PROGRAM prg_Initialise
VAR_INPUT
	ResumeSFC       : BOOL; 		(*	not automatic	*)
	//Added SFC Cycle handle Variables
	
	SFCInit             : BOOL;  //shachar
END_VAR

VAR


(* 8888888888888888   SFC   8888888888888888888888*)
	sCycleName	        : STRING;
	SFCCurrentStep      : STRING;
	SFCErrorPOU         : STRING;
	SFCErrorStep        : STRING;
	SFCError            : BOOL;
	SFCPause            : BOOL;
	
	SFCTipMode          : BOOL;
	SFCTip              : BOOL;
	SFCEnableLimit		: BOOL:=TRUE;
	// Reset Error
	SFCReset			: BOOL;
	ErrorSFC            : BOOL; 	(*	not automatic	*)

	ResetError          : BOOL; 	(*	not automatic	*)
	Last_SFCErrorStep   : STRING; 	(*	not automatic	*)
	//ErrorToPrint        : STRING; 	(*	not automatic	*)
	//Last_ErrorToPrint   : STRING; 	(*	not automatic	*)

 //   stSafety			:ST_BasicCycle;  //shachar
(* 8888888888888888   SFC   8888888888888888888888*)




	Pis             : INT;
	c_PisInitCheck  : INT;
	b_AllPisInitPos : BOOL;

	i               : INT;
	c_LatInitCheck  : INT;

	c_PisResetCleare: INT;

	k               : INT;

	bGeneralDone    : BOOL;
	bPistonDone     : BOOL;
	b_StationDone   : BOOL;
	bLoadConvDone   : BOOL;
	bUnloadConvDone : BOOL;
	bTableDone      : BOOL;
	bStackerDone    : BOOL;
    bManipulatorDone: BOOL;

	init_General    : BOOL;
	init_AllPiston  : BOOL;
	init_AllStation : BOOL;
	init_Table      : BOOL;
	init_LoadConv   : BOOL;
	init_UnloadConv : BOOL;
	init_Stacker    : BOOL;
	init_Manipulator: BOOL;

	bMessLoadInit   : BOOL;
	bMessUnloadInit : BOOL;
	
	sFB_ID          : STRING(4):='004';
	sFB_Num         : STRING(4):='000';
	sActErrorID     : STRING;
	//Added SFC Cycle handle Variables
	fb_SFC_Cycle		    : FB_SFC_Cycle;
	fbFormatString	    	: FB_FORMATSTRING;
	sFullErrorId		    : STRING(12);//sAAAxBBBxEEE
	bReset					: BOOL;

	bIntZoneOk: BOOL;
	bNotPrepare: BOOL;
	p_ManipReset: POINTER TO BOOL;
	p_PowerMotorOn: POINTER TO BOOL;
	p_SafetyStart: POINTER TO BOOL;
   // fbPowerMotorOn			:FB_PowerMotorOn;

	IndexOn: BOOL;
	LoadOn: BOOL;
	UnloadOn: BOOL;
	ManipOn: BOOL;
	p_PowerMotorPower: POINTER TO BOOL;
	p_PowerMotorOff: POINTER TO BOOL;
	iResumeCount: INT;
	iIndexCount: INT;
	iLoadCount: INT;
	iUnloadCount: INT;
	iManipCount: INT;
	p_ManipResume: POINTER TO BOOL;
END_VAR

VAR_IN_OUT
	stOperation	: ST_OperationButtons;	
END_VAR

act_General();
act_Piston();
act_GetErrorID();
fb_SFC_Cycle
( 
	sCycleName:= 'Initialize', 
	bSFCError:= SFCError, 
	sSFCCurrentStep:=SFCCurrentStep , 
	sSFCErrorStep:= SFCErrorStep, 
	sSFCErrorPOU:=SFCErrorPOU , 
	sActErrorID:=sFullErrorId,
	sFB_ModuleDescription:= fb_SFC_Cycle.sCycleName, 
	sLast_SFCErrorStep=>Last_SFCErrorStep , 
	bErrorSFC_Occured=> ErrorSFC, 
	//sErrorToPrint=>ErrorToPrint , 
	//sLast_ErrorToPrint=>Last_ErrorToPrint,
    bSFCInit=>SFCInit , 
	stOperation:= stOperation,
	bResumeSFC:=ResumeSFC , 
	bResetError:=ResetError , 
	bSFCPause:= SFCPause, 
	bResetCycle:=SFCReset
);



IF NOT bStateSafe	
OR init_AllPiston
THEN;
	bGeneralDone:=FALSE;
	bPistonDone:=FALSE;
	b_StationDone:=FALSE;
	bLoadConvDone:=FALSE;
	bUnloadConvDone:=FALSE;
	bTableDone:=FALSE;
	bStackerDone:=FALSE;
	bManipulatorDone:=FALSE;  //shachar
END_IF

ACTION act_General:
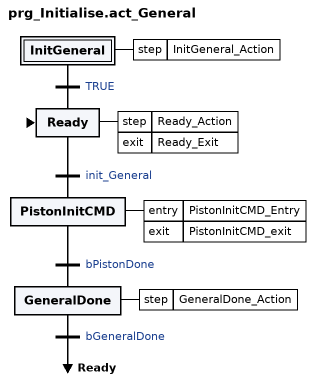
INITIAL_STEP InitGeneral:
    InitGeneral_Action(N);  // step action
END_STEP
TRANSITION FROM InitGeneral TO Ready
    := TRUE;
END_TRANSITION
STEP Ready:
    Ready_Action(N);  // step action
    Ready_Exit(P0);  // exit action
END_STEP
TRANSITION FROM Ready TO PistonInitCMD
    := init_General;
END_TRANSITION
STEP PistonInitCMD:  // min time t#2s
    PistonInitCMD_Entry(P1);  // entry action
    PistonInitCMD_exit(P0);  // exit action
END_STEP
TRANSITION FROM PistonInitCMD TO GeneralDone
    := bPistonDone;
END_TRANSITION
STEP GeneralDone:
    GeneralDone_Action(N);  // step action
END_STEP
TRANSITION FROM GeneralDone TO Ready
    := bGeneralDone;
END_TRANSITION
END_ACTION

ACTION act_GetErrorID:
IF ErrorSFC THEN;
	// Initialization
	IF    Last_SFCErrorStep='WatingForEmergencyOK' 			THEN sActErrorID:='001';
	ELSIF Last_SFCErrorStep='WatingForInterlockOK' 		    THEN sActErrorID:='002';
	ELSIF Last_SFCErrorStep='WatingForMotorsOK' 			THEN sActErrorID:='003';
	ELSIF Last_SFCErrorStep='CheckInitStationDone' 			THEN sActErrorID:='004';
	ELSIF Last_SFCErrorStep='Station_Initialization' 		THEN sActErrorID:='005';
	ELSIF Last_SFCErrorStep='Loader_Initialization' 		THEN sActErrorID:='006';
	ELSIF Last_SFCErrorStep='Unload_Station' 			    THEN sActErrorID:='007';
	ELSIF Last_SFCErrorStep='Measuring_Station' 			THEN sActErrorID:='008';
	ELSIF Last_SFCErrorStep='Gripper_Oriantation' 			THEN sActErrorID:='009';
	ELSIF Last_SFCErrorStep='Index_Homming' 			    THEN sActErrorID:='010';
	ELSIF Last_SFCErrorStep='PaletBypasCheck_1' 			THEN sActErrorID:='011';
	ELSIF Last_SFCErrorStep='PaletCheck_1' 			        THEN sActErrorID:='012';
	ELSIF Last_SFCErrorStep='Cover_Station' 			    THEN sActErrorID:='023';	
	ELSE;
		 sActErrorID:='999';
	END_IF
//ELSIF bWarning THEN;
	// Leave the warning message to print
ELSE;
		 sActErrorID:='000';
END_IF
//*** Error Format ***
fbFormatString(
	sFormat:= '%.3sx%.3sx%.3s', 
	arg1:= F_STRINGEx(sFB_ID), 
	arg2:= F_STRINGEx(sFB_Num), 
	arg3:= F_STRINGEx(sActErrorID), 
	sOut=>sFullErrorId );
	
//(*Clean Last ErrID*)IF NOT SFCPause THEN	sFullErrorId:='';END_IF
END_ACTION

ACTION act_Piston:
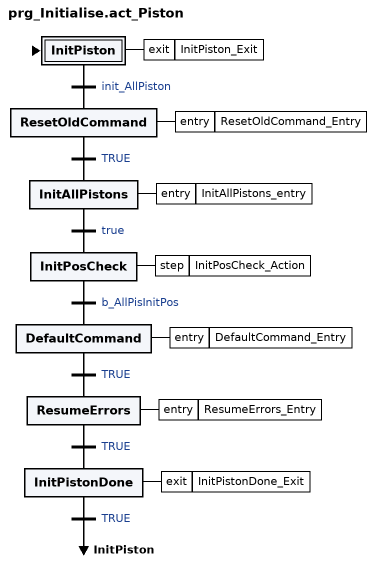
INITIAL_STEP InitPiston:
    InitPiston_Exit(P0);  // exit action
END_STEP
TRANSITION FROM InitPiston TO ResetOldCommand
    := init_AllPiston;
END_TRANSITION
STEP ResetOldCommand:  // min time T#0.1S
    ResetOldCommand_Entry(P1);  // entry action
END_STEP
TRANSITION FROM ResetOldCommand TO InitAllPistons
    := TRUE;
END_TRANSITION
STEP InitAllPistons:  // min time t#1s
    InitAllPistons_entry(P1);  // entry action
END_STEP
TRANSITION FROM InitAllPistons TO InitPosCheck
    := true;
END_TRANSITION
STEP InitPosCheck:
    InitPosCheck_Action(N);  // step action
END_STEP
TRANSITION FROM InitPosCheck TO DefaultCommand
    := b_AllPisInitPos;
END_TRANSITION
STEP DefaultCommand:  // min time T#0.2S
    DefaultCommand_Entry(P1);  // entry action
END_STEP
TRANSITION FROM DefaultCommand TO ResumeErrors
    := TRUE;
END_TRANSITION
STEP ResumeErrors:  // min time T#0.2S
    ResumeErrors_Entry(P1);  // entry action
END_STEP
TRANSITION FROM ResumeErrors TO InitPistonDone
    := TRUE;
END_TRANSITION
STEP InitPistonDone:
    InitPistonDone_Exit(P0);  // exit action
END_STEP
TRANSITION FROM InitPistonDone TO InitPiston
    := TRUE;
END_TRANSITION
END_ACTION

ACTION DefaultCommand_Entry:
	(*FOR Pis:=1 TO 24 BY 1 DO
		db_Lat[Pis].req_DefaultPos:=TRUE;
	END_FOR*)
	
	FOR Pis:=1 TO C_Max_Pistons BY 1 DO
		IF stPis[Pis].b_PistonActive THEN;
			stPis[Pis].req_Init:=TRUE;
		END_IF		
	END_FOR
END_ACTION

ACTION GeneralDone_Action:
init_General:=FALSE;
bGeneralDone:=TRUE;
END_ACTION

ACTION InitAllPistons_entry:
prg_Pistons.bInitAllPiston:=TRUE;
END_ACTION

ACTION InitGeneral_Action:
SFCReset:=FALSE;

init_AllPiston   :=FALSE;
END_ACTION

ACTION InitPiston_Exit:
	b_AllPisInitPos:=FALSE;
	bPistonDone:=FALSE;
END_ACTION

ACTION InitPistonDone_Exit:
	init_AllPiston:=FALSE;
	bPistonDone:=TRUE;
END_ACTION

ACTION InitPosCheck_Action:
			c_PisInitCheck:=0;
	FOR Pis:=1 TO C_Max_Pistons BY 1 DO
		IF fb_Pis[Pis].SFCCurrentStep<>'Ready' AND fb_Pis[Pis].SFCCurrentStep<>''THEN
			c_PisInitCheck:=c_PisInitCheck+1;
		END_IF
	END_FOR

			c_PisResetCleare:=0;
	FOR Pis:=1 TO C_Max_Pistons BY 1 DO
		IF stPis[Pis].b_Reset THEN
			c_PisResetCleare:=c_PisResetCleare+1;
		END_IF
	END_FOR

	(*		c_LatInitCheck:=0;
	FOR Pis:=1 TO 24 BY 1 DO
		IF fb_Lat[Pis].SFCCurrentStep<>'Ready' AND fb_Lat[Pis].SFCCurrentStep<>'' THEN
			c_LatInitCheck:=c_LatInitCheck+1;
		END_IF
	END_FOR*)


		IF 	c_PisInitCheck=0  AND c_LatInitCheck=0 (*AND 	c_PisResetCleare=0*) THEN
			b_AllPisInitPos:=TRUE;
		ELSE
			b_AllPisInitPos:=FALSE;
		END_IF
END_ACTION

ACTION PistonInitCMD_Entry:
init_AllPiston:=TRUE;
END_ACTION

ACTION PistonInitCMD_exit:
Global_Variables.ResumeAll :=TRUE;
END_ACTION

ACTION Ready_Action:
IF TRUE
AND	bPistonDone
(*AND	b_StationDone
AND	bLoadConvDone
AND	bUnloadConvDone
AND	bTableDone
AND (bManipulatorDone OR NOT b_ManipulatorExist)
AND	(bStackerDone OR NOT b_StackerExist)*)
THEN
	bGeneralDone:=TRUE;

ELSE
	bGeneralDone:=FALSE;
END_IF
END_ACTION

ACTION Ready_Exit:
bGeneralDone:=FALSE;
bPistonDone:=FALSE;
b_StationDone:=FALSE;
bLoadConvDone:=FALSE;
bUnloadConvDone:=FALSE;
bTableDone:=FALSE;
bStackerDone:=FALSE;

bManipulatorDone:=FALSE; //shachar
iResumeCount:=0;
END_ACTION

ACTION ResetOldCommand_Entry:
	(*FOR Pis:=1 TO 24 BY 1 DO
		db_Lat[Pis].req_Reset:=TRUE;
	END_FOR*)
	FOR Pis:=1 TO C_Max_Pistons BY 1 DO
		stPis[Pis].b_Reset:=TRUE;
	END_FOR
END_ACTION

ACTION ResumeErrors_Entry:
	(*FOR Pis:=1 TO 24 BY 1 DO
		db_Lat[Pis].req_Resume:=TRUE;
	END_FOR*)
	FOR Pis:=1 TO C_Max_Pistons BY 1 DO
		stPis[Pis].b_Resume:=TRUE;
	END_FOR
END_ACTION

END_PROGRAM

(* stored: Version 1.1.0.1, ProductVersion 3.1.4024.13
   POU prg_Initialise: Id {547dfe07-e15f-49a5-8906-1a326ec23637}, SpecialFunc None
   Folder General: Id {efe61118-d10b-4554-b7e2-cfc68ad8097a}
   Folder Piston: Id {915b62bb-f05b-45db-b566-9bcc993972f9}
   Action act_General: Id {d8f67e11-6dfc-4cdd-b402-56acaf7d55e6}
   Action act_GetErrorID: Id {d06921cf-a63e-4173-a9f9-7618dff90d12}
   Action act_Piston: Id {c1c30121-7ee6-4224-b72d-2c5571419656}
   Action DefaultCommand_Entry: Id {fdc9c316-7914-4767-bd3f-eeabdb22e4ed}
   Action GeneralDone_Action: Id {4ae0d015-5eba-445b-b0a9-b27b0373604b}
   Action InitAllPistons_entry: Id {a53759c3-dcb0-4bf9-85b7-1602b3b3a1ff}
   Action InitGeneral_Action: Id {eaf7217d-7f1e-4ed4-86e4-c1ca1deb192f}
   Action InitPiston_Exit: Id {81262ffa-94cd-4f77-9823-01220b89dabe}
   Action InitPistonDone_Exit: Id {cb2326a3-f022-4764-85dc-08418fc4a3b0}
   Action InitPosCheck_Action: Id {e21c5f29-a93c-4aed-a871-e52f1086b9f9}
   Action PistonInitCMD_Entry: Id {630e0a63-f239-4dbc-8c6a-f04b1ad153af}
   Action PistonInitCMD_exit: Id {64c55cf3-63af-406c-b170-3461aabacc57}
   Action Ready_Action: Id {92f1df72-5324-423e-8850-d013024f6f59}
   Action Ready_Exit: Id {60c681e3-4bcf-4070-ae7f-84b907b0ee02}
   Action ResetOldCommand_Entry: Id {6847173e-ff86-4ed0-a862-24256ccb17c1}
   Action ResumeErrors_Entry: Id {655a0cf4-61f8-4a22-8784-f3b9adc39cbe} *)
